TYPE ST_Halytykset :
STRUCT
	nID:				LINT;
	tAikaleima:			DATE_AND_TIME;
	sKoodi:				STRING(50);	
	sKuvaus:			STRING(255);

	
END_STRUCT
END_TYPE

(* stored: Version 1.1.0.1
   DUT ST_Halytykset: Id {9a263320-f20b-417d-a0f2-392ebf9d0608} *)
